# B&R Automation Studio project DriveControl
Automation Studio 4.5.2.102; Default project; technology packages: Acp10Arnc0 5.2.1

## Configuration SampleText

CPU 4PP065.0571-P74, AutomationRuntime D4.52, Build 4.1.2, Vc V4.25.0, Safety 1.6

### Task classes (Cpu.sw)
```
Cyclic#1 (cycle 2000 us, tolerance 0 us):
  ncsdcctrl <- ncsdcctrl.prg
Cyclic#4:
  Program <- Program.prg
NcDataObjects: acp10etxen <- acp10etxen.dob, gAxis01a <- gAxis01obj.gAxis01a.dob, gAxis01i <- gAxis01obj.gAxis01i.dob
Libraries: Acp10sdc, sys_lib, Runtime, asstring, Acp10man, Acp10par, NcGlobal, Acp10_MC, brsystem, AsBrStr, Library
```

### Hardware
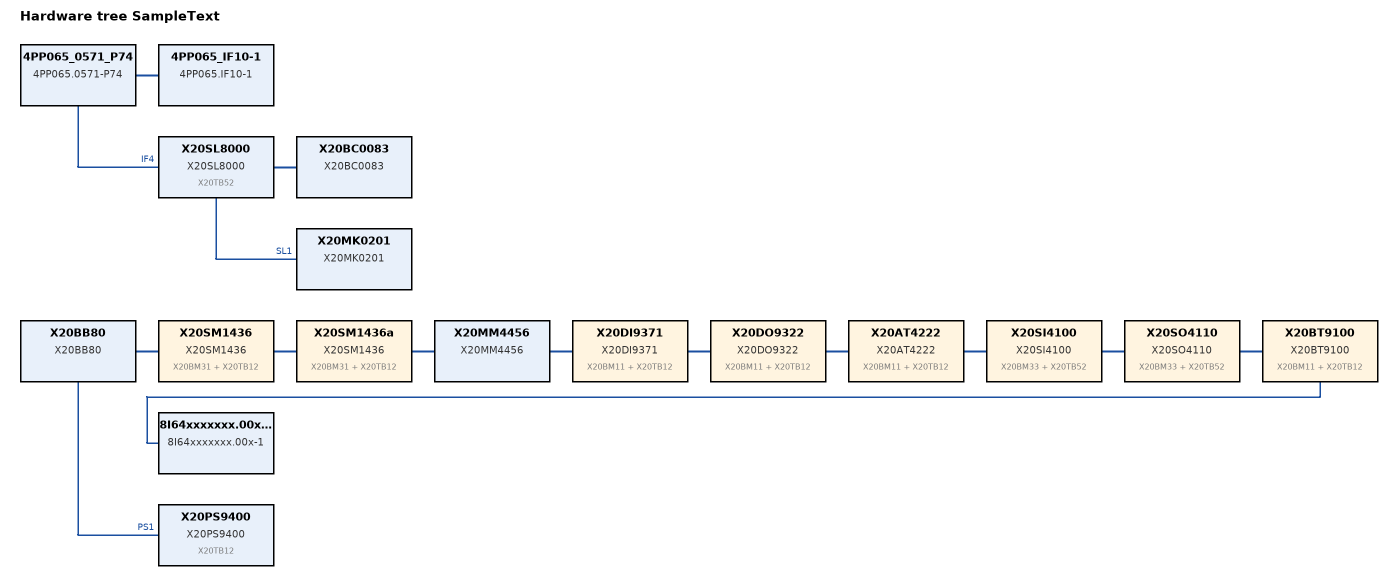
```
4PP065_0571_P74 : 4PP065.0571-P74 v1.1.2.0
  Connector IF5:
    ActivateDevice = 1
    Mode = Manual
    InternetAddress = 10.0.1.10
    SubnetMask = 255.255.255.0
  ConfigurationID = labBR
  TimerDeviceType = EPLX2X
  TimerDevice = 4PP065_0571_P74.IF4
  TaskClassIdleTime = 2000
  Cyclic1Duration = 2000
  Cyclic1Tolerance = 0
  Cyclic1Output = 1
4PP065_IF10-1 : 4PP065.IF10-1 v1.0.3.0  [SS -> 4PP065_0571_P74.SS1]
8I64xxxxxxx.00x-1 : 8I64xxxxxxx.00x-1 v1.3.9.1  [X2X1 -> X20BT9100.X2X1 [Cable Type=X2XCable, Length=10, Version=1.0.0.2]]
  packedETAD = packed
  packedETI = packed
  packedCMDD = packed
  packedCMI = packed
  ACC = 30
  DEC = 30
  UNS = 220
  NCR = 10
  NSP = 890
  COS = 64
  RSC = 33000
X20AT4222 : X20AT4222 v1.2.3.0  [SS1 -> X20TB12e.SS; SL -> X20BM11c.SL1]
X20BB80 : X20BB80 v1.0.2.0
X20BC0083 : X20BC0083 v2.9.0.0  [PLK1 -> X20SL8000.PLK2 (NodeNumber=2) [Cable Type=PowerlinkCable, Length=10, Version=1.0.0.2]; SL -> X20BB80.SL1]
X20BM11 : X20BM11 v1.0.0.1  [X2X1 -> X20BM33a.X2X2]
X20BM11a : X20BM11 v1.0.0.1  [X2X1 -> X20MM4456.X2X2]
X20BM11b : X20BM11 v1.0.0.1  [X2X1 -> X20BM11a.X2X2]
X20BM11c : X20BM11 v1.0.0.1  [X2X1 -> X20BM11b.X2X2]
X20BM31 : X20BM31 v1.0.0.1  [X2X1 -> X20BB80.IF1]
X20BM31a : X20BM31 v1.0.0.1  [X2X1 -> X20BM31.X2X2]
X20BM33 : X20BM33 v1.0.0.4  [X2X1 -> X20BM11c.X2X2]
X20BM33a : X20BM33 v1.0.0.4  [X2X1 -> X20BM33.X2X2]
X20BT9100 : X20BT9100 v1.0.3.0  [SS1 -> X20TB12f.SS; SL -> X20BM11.SL1]
X20DI9371 : X20DI9371 v1.0.2.0  [SS1 -> X20TB12c.SS; SL -> X20BM11a.SL1]
X20DO9322 : X20DO9322 v1.0.3.0  [SS1 -> X20TB12d.SS; SL -> X20BM11b.SL1]
X20MK0201 : X20MK0201 v1.0.0.0  [SL -> X20SL8000.SL1]
X20MM4456 : X20MM4456 v1.1.5.0  [X2X1 -> X20BM31a.X2X2]
X20PS9400 : X20PS9400 v1.0.2.4  [SS1 -> X20TB12.SS; PS -> X20BB80.PS1]
X20SI4100 : X20SI4100 v1.10.1.1  [SS1 -> X20TB52.SS; SL -> X20BM33.SL1]
X20SL8000 : X20SL8000 v1.6.5.1  [PLK1 -> 4PP065_0571_P74.IF4 (NodeNumber=1) [Cable Type=PowerlinkCable, Length=10, Version=1.0.0.2]; PLK2 -> X20BC0083.PLK1 (NodeNumber=1) [Cable Type=PowerlinkCable, Length=10, Version=1.0.0.2]; SS1 -> X20TB52b.SS]
  SafeProject = SafeLOGIC-1
X20SM1436 : X20SM1436 v2.3.0.0  [SS1 -> X20TB12a.SS; SL -> X20BM31.SL1]
X20SM1436a : X20SM1436 v2.3.0.0  [SS1 -> X20TB12b.SS; SL -> X20BM31a.SL1]
X20SO4110 : X20SO4110 v1.10.1.1  [SS1 -> X20TB52a.SS; SL -> X20BM33a.SL1]
  SafeModuleID = 3
X20TB12 : X20TB12 v1.0.0.0
X20TB12a : X20TB12 v1.0.0.0
X20TB12b : X20TB12 v1.0.0.0
X20TB12c : X20TB12 v1.0.0.0
X20TB12d : X20TB12 v1.0.0.0
X20TB12e : X20TB12 v1.0.0.0
X20TB12f : X20TB12 v1.0.0.0
X20TB52 : X20TB52 v1.0.0.1
X20TB52a : X20TB52 v1.0.0.1
X20TB52b : X20TB52 v1.0.0.1
```

### IoMap.iom - 4PP065_0571_P74/IoMap.iom
```iecst
VAR_CONFIG
	Cyclic#1.gAxis01_DrvIf.iLifeCnt AT %IB."8I64xxxxxxx.00x-1".SDC_LifeCnt;
	Cyclic#1.gAxis01_DrvIf.iDrvOK AT %IX."8I64xxxxxxx.00x-1".ETAD_Input_Bool_02;
	Cyclic#1.gAxis01_DrvIf.oSetTime AT %QW."8I64xxxxxxx.00x-1".SDC_SetTime;
	Cyclic#1.::stateMachine.speed AT %QW."8I64xxxxxxx.00x-1".LFRD_Output;
	Cyclic#1.gAxis01_DiDoIf.iLifeCntDriveReady AT %IB."8I64xxxxxxx.00x-1".SDC_LifeCnt;
	Cyclic#1.gAxis01_DiDoIf.iLifeCntDriveEnable AT %IB."8I64xxxxxxx.00x-1".SDC_LifeCnt;
	Cyclic#1.gAxis01_DiDoIf.oDriveEnable AT %QX."8I64xxxxxxx.00x-1".CMDD_Output_Bool_00;
	Cyclic#1.gAxis01_ModuleOk AT %QX."8I64xxxxxxx.00x-1".CMDD_Output_Bool_01;
	Cyclic#1.gAxis01_ModuleOk AT %QX."8I64xxxxxxx.00x-1".CMDD_Output_Bool_02;
	Cyclic#1.gAxis01_ModuleOk AT %IX."8I64xxxxxxx.00x-1".ModuleOk;
	Cyclic#1.gAxis01_DiDoIf.oDriveEnable AT %QX."8I64xxxxxxx.00x-1".CMDD_Output_Bool_03;
	Cyclic#1.gAxis01_DiDoIf.iDriveReady AT %IX."8I64xxxxxxx.00x-1".ETAD_Input_Bool_02;
	::stateMachine.state AT %IW."8I64xxxxxxx.00x-1".ETAD_Input;
	::stateMachine.command AT %QW."8I64xxxxxxx.00x-1".CMDD_Output;
	::doorSM.direction AT %IX."X20DI9371".DigitalInput01;
	::doorSM.sw1 AT %IX."X20DI9371".DigitalInput02;
	::doorSM.sw2 AT %IX."X20DI9371".DigitalInput03;
	::doorSM.sw3 AT %IX."X20DI9371".DigitalInput04;
	::doorSM.sw4 AT %IX."X20DI9371".DigitalInput05;
	::ledSM.led1 AT %QX."X20DO9322".DigitalOutput02;
	::ledSM.led2 AT %QX."X20DO9322".DigitalOutput03;
	::ledSM.led3 AT %QX."X20DO9322".DigitalOutput04;
	::ledSM.led4 AT %QX."X20DO9322".DigitalOutput05;
END_VAR
```

### Acp10cfg.ncc - 4PP065_0571_P74/Motion/Acp10cfg.ncc
```
NcConfiguration (Version=5.02.1, NcSwId=Acp10)
  ACP10CF1_typ:
    cnt_nettrc_rec_drive = 1500
    bufsize_trace_upload = 1200
    tc_nc_man_task = Cyclic #1
    glob_pv_as_ncobject = Yes
    ncsys_dl_broadcast = Yes
    ncsys_dl_acp_reset = Yes
    safemc_log_err_to_ax = Yes
    network_init:
      ncsw_init_execute = Yes
      automatic_execute = No
      node_nr_warning = Yes
      net_err_before_ncact = Yes
    nettrc:
      enter_parsecrec = Yes
      enter_ncaction = Yes
      save_ring_startidx = Yes
    cam_prof_download:
      cam_dat_dl_parallel = No
      tc_cam_dl_parallel = Task class for NC Manager task
    sdc_if[0]:
      if_name = SDC_IF1
      mc_broadcast_size = 800
      mc_broadcast_extdat = No
```

### Acp10map.ncm - 4PP065_0571_P74/Motion/Acp10map.ncm
```
NcMapping (NcSwId=Acp10)
  NcObject gAxis01 (ModuleId=8I64xxxxxxx.00x-1, ModuleAddress=SDC_IF1.ST1, Type=ncAXIS, Channel=1, AcoposSimulation=Off, InitParameter=gAxis01i, AcoposParameter=gAxis01a, Disabled=FALSE, ModuleDisabled=FALSE)
```

- Physical/SampleText/4PP065_0571_P74/PvMap.vvm: same as Physical/SampleText/4PP065_0571_P74/Cpu.per
## Configuration Simulation

CPU , AutomationRuntime J4.25

### Task classes (Cpu.sw)
```
Libraries: AsIecCon, astime
```

### Hardware
```
PC_any : PC_any v1.1.0.0 (OrderNumber=PC)
```

- Physical/Simulation/PC_any/Cpu.per: same as Physical/SampleText/4PP065_0571_P74/Cpu.per
- Physical/Simulation/PC_any/PvMap.vvm: same as Physical/Simulation/PC_any/IOMap.iom
## Logical view

Binary libraries used (declarations not repeated): RUNTIME, OPERATOR, AsIecCon, astime, sys_lib, asstring, Acp10man 5.02.1, Acp10par 5.02.1, NcGlobal 5.02.1, Acp10sdc 5.02.1, Acp10_MC 5.02.1, brsystem, AsBrStr

### Global.var - Global variables
```iecst
VAR
	gAxis01 : ACP10AXIS_typ := (0);
	gAxis01_HW : SdcHwCfg_typ := (0);
	gAxis01_DrvIf : SdcDrvIf16_typ := (0);
	gAxis01_DiDoIf : SdcDiDoIf_typ := (0);
	gAxis01_ModuleOk : BOOL := 0;
	doorSM : DoorStateMashine := (0);
	driveSM : DriveStateMashine := (0);
	ledSM : LedStateMashine := (0);
	stateMachine : DriveStateMashine := (0);
END_VAR
```


### Program Logical/ncsdcctrl (IEC)

#### ncsdcctrlCyclic.st
```iecst
PROGRAM _CYCLIC

(* ### BEGIN gAxis01 ### *)

(* life counter emulation of digital inputs *)
        gAxis01_DiDoIf.iLifeCntReference := gAxis01_DiDoIf.iLifeCntReference + 1;
        gAxis01_DiDoIf.iLifeCntNegHwEnd  := gAxis01_DiDoIf.iLifeCntNegHwEnd  + 1;
        gAxis01_DiDoIf.iLifeCntPosHwEnd  := gAxis01_DiDoIf.iLifeCntPosHwEnd  + 1;

(* ### END gAxis01 ### *)

END_PROGRAM
```

#### ncsdcctrlInit.st
```iecst
PROGRAM _INIT

(* ### BEGIN gAxis01 ### *)

(* initialize variables *)
        gAxis01_HW.DrvIf_Typ := ncSDC_DRVSERVO16;
        brsstrcpy(ADR(gAxis01_HW.DrvIf_Name[0]), ADR('gAxis01_DrvIf'));
        gAxis01_HW.DiDoIf_Typ := ncSDC_DIDO;
        brsstrcpy(ADR(gAxis01_HW.DiDoIf_Name[0]), ADR('gAxis01_DiDoIf'));

(* force variable offset generation *)
        gAxis01.size                      := gAxis01.size;
        gAxis01_DrvIf.iLifeCnt            := gAxis01_DrvIf.iLifeCnt;
        gAxis01_DiDoIf.iLifeCntDriveReady := gAxis01_DiDoIf.iLifeCntDriveReady;
        gAxis01_ModuleOk                  := gAxis01_ModuleOk;

(* assign your hardware inputs here*)

(*      gAxis01_DiDoIf.iPosHwEnd  := gAxis01_DiDoIf.iPosHwEnd;
        gAxis01_DiDoIf.iNegHwEnd  := gAxis01_DiDoIf.iNegHwEnd;
        gAxis01_DiDoIf.iReference := gAxis01_DiDoIf.iReference;
 *)

(* ### END gAxis01 ### *)

END_PROGRAM
```

### Data object Logical/acp10etxen (Ett)

- acp10etxen.ett (not shown)

### Package Logical/gAxis01obj - gAxis01obj

### Data object Logical/gAxis01obj/gAxis01a (Apt)

#### gAxis01a.apt
```
AcoposParameterTable:
  Root Parameters:
    230 = PCTRL_S_SET (Name=PCTRL_S_ACT_PARID)
    64201 = 546116.666666667 (Name=SERVO_V_MAX_OUTPUT)
```

### Data object Logical/gAxis01obj/gAxis01i (Ax)

#### gAxis01i.ax
```
InitParameter (Version=5.2.1, NcSwId=Acp10)
  ACP10AXIS_typ:
    dig_in:
      level:
        reference = ncACTIV_HI
        pos_hw_end = ncACTIV_LO
        neg_hw_end = ncACTIV_LO
        trigger1 = ncACTIV_HI
        trigger2 = ncACTIV_LO + ncQUICKSTOP
    encoder_if:
      parameter:
        count_dir = ncSTANDARD
        scaling:
          load:
            units = 1000
            rev_motor = 1
    limit:
      parameter:
        v_pos = 10000
        v_neg = 10000
        a1_pos = 50000
        a2_pos = 50000
        a1_neg = 50000
        a2_neg = 50000
        t_jolt = 0
        t_in_pos = 0
        pos_sw_end = 2000000000
        neg_sw_end = -2000000000
        ds_warning = 500
        ds_stop = 1000
        a_stop = 1.0e30
        dv_stop = 0
        dv_stop_mode = ncOFF
    controller:
      mode = ncPOSITION
      position:
        kv = 50
        tn = 0
        t_predict = 0.01
        t_total = 0.01
        p_max = 1.0e30
        i_max = 0
      speed:
        kv = 2.0
        tn = 0
        t_filter = 0.0
        isq_filter1:
          type = ncOFF
          a0 = 0.0
          a1 = 0.0
          b0 = 0.0
          b1 = 0.0
          b2 = 0.0
          c0_par_id = 0
          c1_par_id = 0
        isq_filter2:
          type = ncOFF
          a0 = 0.0
          a1 = 0.0
          b0 = 0.0
          b1 = 0.0
          b2 = 0.0
          c0_par_id = 0
          c1_par_id = 0
        isq_filter3:
          type = ncOFF
          a0 = 0.0
          a1 = 0.0
          b0 = 0.0
          b1 = 0.0
          b2 = 0.0
          c0_par_id = 0
          c1_par_id = 0
      uf:
        type = ncLINEAR + ncCORRECTION
        auto_config = ncMOTOR_PAR
        u0 = 0
        un = 0
        fn = 50.0
        k_f_slip = 0
      ff:
        torque_load = 0.0
        torque_pos = 0.0
        torque_neg = 0.0
        kv_torque = 0.0
        inertia = 0.0
        t_filter_a = 0.0
    move:
      stop:
        parameter[0]:
          decel_ramp = ncA_LIMIT
          controller = ncON
        parameter[1]:
          decel_ramp = ncA_LIMIT
          controller = ncON
        parameter[2]:
          decel_ramp = ncA_LIMIT
          controller = ncON
        parameter[3]:
          decel_ramp = ncA_LIMIT
          controller = ncON
        quickstop:
          decel_ramp = ncA_LIMIT
          t_jolt = 0
        drive_error:
          decel_ramp = ncA_LIMIT
      homing:
        parameter:
          s = 0
          v_switch = 5000
          v_trigger = 500
          a = 50000
          mode = ncDIRECT
          edge_sw = ncPOSITIVE
          start_dir = ncPOSITIVE
          trigg_dir = ncPOSITIVE
          ref_pulse = ncOFF
          fix_dir = ncOFF
          tr_s_block = 0
          torque_lim = 0
          ds_block = 0
          ds_stop = 0
      basis:
        parameter:
          v_pos = 5000
          v_neg = 5000
          a1_pos = 50000
          a2_pos = 50000
          a1_neg = 50000
          a2_neg = 50000
    message:
      text:
        parameter:
          format = ncBREAK
          columns = 80
          data_modul = acp10etxen
```

### Library Logical/Library (ANSIC)

#### Types.typ - Exported data types
```iecst
TYPE
	DoorStates :
		(
		ST_INIT,
		ST_UNKNOWN,
		ST_OPEN,
		ST_CLOSE,
		ST_ACC_POS,
		ST_ACC_NEG,
		ST_POS,
		ST_NEG,
		ST_DEC_POS,
		ST_DEC_NEG
		);
END_TYPE
```

#### Constants.var - Exported constants
```iecst
VAR CONSTANT
	SPEED_SLOW : INT := 300; (*Slow speed: S0-S1, S2-S3, position search*)
	SPEED_FAST : INT := 800; (*Fast speed: S1-S2*)
	SPEED_STOP : INT := 0;
	DRV_STATE_MASK : UINT := 16#006F; (*Status word mask*)
	STATE_SWITCHED_ON : UINT := 16#0021; (*Ready to switch on*)
	STATE_READY : UINT := 16#0023; (*Switched on*)
	STATE_ENABLED : UINT := 16#0027; (*Operation enabled*)
	STATE_FAULT_BIT : UINT := 16#0008; (*Fault bit*)
	CMD_SHUTDOWN : UINT := 16#0006;
	CMD_SWITCH_ON : UINT := 16#0007;
	CMD_ENABLE : UINT := 16#000F;
	CMD_FAULT_RESET : UINT := 16#0080;
	BLINK_HALF_PERIOD_MS : UDINT := 500; (*1 Hz blink*)
END_VAR
```

#### Library.fun - Exported functions and function blocks
```iecst
{REDUND_ERROR} FUNCTION_BLOCK DriveStateMashine (*Frequency inverter control (CiA402)*) (*$GROUP=User,$CAT=User,$GROUPICON=User.png,$CATICON=User.png*)
	VAR_INPUT
		state : UINT; (*Inverter status word (ETAD)*)
		enable : BOOL; (*Enable FB*)
		speedSet : INT; (*Speed setpoint from door logic*)
	END_VAR
	VAR_OUTPUT
		command : UINT; (*Inverter control word (CMDD)*)
		speed : INT; (*Speed to inverter (LFRD)*)
	END_VAR
END_FUNCTION_BLOCK

{REDUND_ERROR} FUNCTION_BLOCK DoorStateMashine (*Door state machine*) (*$GROUP=User,$CAT=User,$GROUPICON=User.png,$CATICON=User.png*)
	VAR_INPUT
		state : UINT; (*Inverter status word*)
		sw1 : BOOL; (*S0 - door open*)
		sw2 : BOOL; (*S1*)
		sw3 : BOOL; (*S2*)
		sw4 : BOOL; (*S3 - door closed*)
		direction : BOOL; (*Switch: 1 - close, 0 - open*)
	END_VAR
	VAR_OUTPUT
		speed : INT; (*Speed setpoint*)
		doorState : DoorStates; (*Current door state*)
	END_VAR
	VAR
		s0Prev : BOOL; (*Sensor levels on previous cycle*)
		s1Prev : BOOL;
		s2Prev : BOOL;
		s3Prev : BOOL;
	END_VAR
END_FUNCTION_BLOCK

{REDUND_ERROR} FUNCTION_BLOCK LedStateMashine (*LED indication*) (*$GROUP=User,$CAT=User,$GROUPICON=User.png,$CATICON=User.png*)
	VAR_INPUT
		state : UINT; (*Door state*)
		cycleTime : UDINT; (*Task cycle time, ms*)
	END_VAR
	VAR_OUTPUT
		led1 : BOOL; (*S0*)
		led2 : BOOL; (*S1*)
		led3 : BOOL; (*S2*)
		led4 : BOOL; (*S3*)
		timer : INT; (*Blink timer, ms*)
	END_VAR
	VAR
		elapsed : UDINT;
		blink : BOOL;
	END_VAR
END_FUNCTION_BLOCK
```

#### DriveStateMashine.c
```c
#include <bur/plctypes.h>
#ifdef __cplusplus
	extern "C"
	{
#endif
#include "Library.h"
#ifdef __cplusplus
	};
#endif

/*
 * Управление частотным преобразователем (рис. 2.9, профиль CiA 402 / DRIVECOM).
 * state   - слово состояния ETAD, анализируется по маске 0x6F
 * command - слово управления CMDD
 * speed   - задание скорости LFRD (выдаётся только в состоянии "работа разрешена")
 */
void DriveStateMashine(struct DriveStateMashine* inst)
{
	UINT st = inst->state & DRV_STATE_MASK;

	/* Работа блока запрещена -> SHUTDOWN, скорость 0 */
	if (!inst->enable)
	{
		inst->command = CMD_SHUTDOWN;
		inst->speed   = 0;
		return;
	}

	/* Авария ПЧ -> сброс ошибки */
	if (inst->state & STATE_FAULT_BIT)
	{
		inst->command = CMD_FAULT_RESET;
		inst->speed   = 0;
		return;
	}

	if (st == STATE_ENABLED)
	{
		/* Работа разрешена - передаём задание скорости */
		inst->command = CMD_ENABLE;
		inst->speed   = inst->speedSet;
	}
	else if (st == STATE_READY)
	{
		/* SWITCHED ON -> разрешить работу */
		inst->command = CMD_ENABLE;
		inst->speed   = 0;
	}
	else if (st == STATE_SWITCHED_ON)
	{
		/* READY TO SWITCH ON -> включить */
		inst->command = CMD_SWITCH_ON;
		inst->speed   = 0;
	}
	else
	{
		/* DISABLED (switch on disabled) и прочие -> SHUTDOWN */
		inst->command = CMD_SHUTDOWN;
		inst->speed   = 0;
	}
}
```

#### DoorStateMashine.c
```c
#include <bur/plctypes.h>
#ifdef __cplusplus
	extern "C"
	{
#endif
	#include "Library.h"
#ifdef __cplusplus
	};
#endif

/*
 * Конечный автомат защитной двери (рис. 2.6, 2.11).
 *
 * Датчики:  sw1 = S0 (дверь открыта), sw2 = S1, sw3 = S2, sw4 = S3 (дверь закрыта)
 * Тумблер:  direction = 1 - закрыть (движение S0 -> S3, скорость > 0, состояния *_POS)
 *           direction = 0 - открыть (движение S3 -> S0, скорость < 0, состояния *_NEG)
 * Скорость: S0-S1 и S2-S3 - SPEED_SLOW, S1-S2 - SPEED_FAST.
 *
 * Переходы по датчикам выполняются по ИЗМЕНЕНИЮ логического уровня
 * (0 -> 1 или 1 -> 0), а не по самому значению. Для этого блок хранит
 * уровни датчиков с прошлого цикла (s0Prev..s3Prev).
 * Это относится ко всем датчикам, включая концевые S0 и S3.
 * Тумблер direction работает по уровню - он задаёт, куда ехать.
 *
 * Переходы только последовательные (рис. 2.11): каждый датчик проверяется
 * лишь в том состоянии, которое заканчивается на нём. Перескочить через
 * состояние нельзя. Реверс тумблером - только на тот же отрезок хода
 * (ACC_POS <-> DEC_NEG, POS <-> NEG, DEC_POS <-> ACC_NEG).
 */
void DoorStateMashine(struct DoorStateMashine* inst)
{
	/* Текущие уровни датчиков */
	BOOL s0 = inst->sw1;
	BOOL s1 = inst->sw2;
	BOOL s2 = inst->sw3;
	BOOL s3 = inst->sw4;

	/* Изменение уровня относительно прошлого цикла */
	BOOL s0Changed = (s0 != inst->s0Prev);
	BOOL s1Changed = (s1 != inst->s1Prev);
	BOOL s2Changed = (s2 != inst->s2Prev);
	BOOL s3Changed = (s3 != inst->s3Prev);

	BOOL driveOn = ((inst->state & DRV_STATE_MASK) == STATE_ENABLED);
	DoorStates stateAtStart;

	/* Пропал ПЧ (авария/выключение) - всё заново, через поиск положения */
	if (!driveOn && inst->doorState != ST_INIT)
		inst->doorState = ST_INIT;

	stateAtStart = inst->doorState;

	switch (inst->doorState)
	{
		case ST_INIT:          /* ожидание включения ПЧ */
			inst->speed = SPEED_STOP;
			if (driveOn)
				inst->doorState = ST_UNKNOWN;
			break;

		case ST_UNKNOWN:       /* поиск положения: медленно в сторону тумблера */
			inst->speed = inst->direction ? SPEED_SLOW : -SPEED_SLOW;
			if (!inst->direction && s0Changed)
				inst->doorState = ST_OPEN;
			else if (inst->direction && s3Changed)
				inst->doorState = ST_CLOSE;
			break;

		case ST_OPEN:          /* стоим в S0 */
			inst->speed = SPEED_STOP;
			if (inst->direction)
				inst->doorState = ST_ACC_POS;
			break;

		case ST_ACC_POS:       /* S0 -> S1, медленно */
			inst->speed = SPEED_SLOW;
			if (!inst->direction)
				inst->doorState = ST_DEC_NEG;      /* реверс: назад к S0 */
			else if (s1Changed)
				inst->doorState = ST_POS;
			break;

		case ST_POS:           /* S1 -> S2, быстро */
			inst->speed = SPEED_FAST;
			if (!inst->direction)
				inst->doorState = ST_NEG;
			else if (s2Changed)
				inst->doorState = ST_DEC_POS;
			break;

		case ST_DEC_POS:       /* S2 -> S3, медленно */
			inst->speed = SPEED_SLOW;
			if (!inst->direction)
				inst->doorState = ST_ACC_NEG;
			else if (s3Changed)
				inst->doorState = ST_CLOSE;
			break;

		case ST_CLOSE:         /* стоим в S3 */
			inst->speed = SPEED_STOP;
			if (!inst->direction)
				inst->doorState = ST_ACC_NEG;
			break;

		case ST_ACC_NEG:       /* S3 -> S2, медленно */
			inst->speed = -SPEED_SLOW;
			if (inst->direction)
				inst->doorState = ST_DEC_POS;      /* реверс: назад к S3 */
			else if (s2Changed)
				inst->doorState = ST_NEG;
			break;

		case ST_NEG:           /* S2 -> S1, быстро */
			inst->speed = -SPEED_FAST;
			if (inst->direction)
				inst->doorState = ST_POS;
			else if (s1Changed)
				inst->doorState = ST_DEC_NEG;
			break;

		case ST_DEC_NEG:       /* S1 -> S0, медленно */
			inst->speed = -SPEED_SLOW;
			if (inst->direction)
				inst->doorState = ST_ACC_POS;
			else if (s0Changed)
				inst->doorState = ST_OPEN;
			break;

		default:
			inst->speed = SPEED_STOP;
			inst->doorState = ST_INIT;
			break;
	}

	/* Запоминаем уровни для следующего цикла.
	   Пока ждём ПЧ (ST_INIT), держим "прошлые" уровни равными 0:
	   если дверь уже стоит на датчике, при входе в ST_UNKNOWN
	   это будет воспринято как изменение уровня 0 -> 1. */
	if (stateAtStart == ST_INIT || inst->doorState == ST_INIT)
	{
		inst->s0Prev = 0;
		inst->s1Prev = 0;
		inst->s2Prev = 0;
		inst->s3Prev = 0;
	}
	else
	{
		inst->s0Prev = s0;
		inst->s1Prev = s1;
		inst->s2Prev = s2;
		inst->s3Prev = s3;
	}
}
```

#### LedStateMashine.c
```c
#include <bur/plctypes.h>
#ifdef __cplusplus
	extern "C"
	{
#endif
	#include "Library.h"
#ifdef __cplusplus
	};
#endif

/*
 * Индикация положения двери (рис. 2.11).
 * state - состояние двери (DoorStates), led1..led4 -> индикаторы S0..S3.
 * В ST_UNKNOWN все индикаторы мигают с частотой 1 Гц (500 мс горят / 500 мс нет).
 * cycleTime - время цикла задачи в мс (передаётся из программы, см. Main.c).
 * timer - текущее время внутри полупериода мигания, мс.
 */
static void SetLeds(struct LedStateMashine* inst, BOOL l1, BOOL l2, BOOL l3, BOOL l4)
{
	inst->led1 = l1;
	inst->led2 = l2;
	inst->led3 = l3;
	inst->led4 = l4;
}

void LedStateMashine(struct LedStateMashine* inst)
{
	UDINT dt = inst->cycleTime;
	if (dt == 0)
		dt = 100;   /* на случай, если время цикла не задано */

	switch (inst->state)
	{
		case ST_UNKNOWN:
			inst->elapsed += dt;
			if (inst->elapsed >= BLINK_HALF_PERIOD_MS)
			{
				inst->elapsed = 0;
				inst->blink = !inst->blink;
			}
			SetLeds(inst, inst->blink, inst->blink, inst->blink, inst->blink);
			break;

		case ST_OPEN:     SetLeds(inst, 0, 0, 0, 0); break;
		case ST_ACC_POS:  SetLeds(inst, 1, 0, 0, 0); break;
		case ST_POS:      SetLeds(inst, 1, 1, 0, 0); break;
		case ST_DEC_POS:  SetLeds(inst, 1, 1, 1, 0); break;
		case ST_CLOSE:    SetLeds(inst, 1, 1, 1, 1); break;
		case ST_ACC_NEG:  SetLeds(inst, 1, 1, 1, 0); break;
		case ST_NEG:      SetLeds(inst, 1, 1, 0, 0); break;
		case ST_DEC_NEG:  SetLeds(inst, 1, 0, 0, 0); break;

		case ST_INIT:
		default:
			SetLeds(inst, 0, 0, 0, 0);
			break;
	}

	if (inst->state != ST_UNKNOWN)
	{
		inst->elapsed = 0;
		inst->blink = 0;
	}
	inst->timer = (INT)inst->elapsed;
}
```

### Program Logical/Program (ANSIC)

#### Main.c - Init, cyclic, exit code
```c
#include <bur/plctypes.h>

#ifdef _DEFAULT_INCLUDES
	#include <AsDefault.h>
#endif

void _INIT ProgramInit(void)
{
	stateMachine.enable   = 0;
	stateMachine.speedSet = 0;
	stateMachine.command  = CMD_SHUTDOWN;
	stateMachine.speed    = 0;

	doorSM.doorState = ST_INIT;
	doorSM.speed     = 0;

	ledSM.state = ST_INIT;
	ledSM.led1  = 0;
	ledSM.led2  = 0;
	ledSM.led3  = 0;
	ledSM.led4  = 0;
}

void _CYCLIC ProgramCyclic(void)
{
	/* 1. Логика двери: датчики и тумблер приходят через мэпинг*/
	doorSM.state = stateMachine.state;
	DoorStateMashine(&doorSM);

	/* 2. Управление частотным преобразователем */
	stateMachine.enable   = 1;
	stateMachine.speedSet = doorSM.speed;
	DriveStateMashine(&stateMachine);

	/* 3. Индикация положения двери */
	ledSM.state = (UINT)doorSM.doorState;
	LedStateMashine(&ledSM);
}

void _EXIT ProgramExit(void)
{

}
```
